Fanuc KAREL source: KT00228.KL

PROGRAM KT00228
%NOLOCKGROUP
VAR
  B1: BOOLEAN
  I2: INTEGER
  OUT: INTEGER
BEGIN
  B1 = TRUE
    I2 = 3
  OUT = B1 OR I2
END KT00228
